FUNCTION_BLOCK FB_Gr00Utility
(*

The function block used to control general utility of the machine.

Constructor: 		Patryk Panylo
Company:		E. Riexinger GmbH
Date:			28.04.2015
Version:			1.00

Date:			Revision:		Who:				Comment
dd.mm.yyyy		x.xx			Initials			comment

*)
VAR_INPUT
	(* Input variables / Eingang Variablen *)
	bSignalStart					:BOOL;						(* Signal "Start" / Signal "Start" *)
	bSignalStop					:BOOL;						(* Signal "Stop" / Signal "Stop" *)
	bSignalAbort					:BOOL;						(* Signal "Abort" / Signal "Abort" *)
	bSignalHome					:BOOL;						(* Signal "Home" / Signal "Grundstellung" *)
	bSignalReference				:BOOL;						(* Signal "Reference" / Signal "Referenz" *)
	bSignalReset					:BOOL;						(* Signal "Reset" / Signal "Reset *)
	bSignalMachinePurge			:BOOL;						(* Machine purge *)
	bAutoStartRelease			:BOOL;						(* Auto start release *)
	bHomeStartRelease			:BOOL;						(* Home start release *)
	bAutoToHome				:BOOL;						(* If auto completed go to home *)
	bHomeCompleted				:BOOL;						(* Home completed signal *)
	bAutoCompleted				:BOOL;						(* Auto completed signal *)
	bAllDoorsClosed 				:BOOL;						(* All doors closed *)
	bAllDoorsLocked 				:BOOL;						(* All doors locked *)
	bLightCurtainOk				:BOOL;						(* Light curtain ok *)
	bExeCounter					:BOOL;						(* Execute counter *)
	bResetCounterUser			:BOOL;						(* Reset counter user *)
	bStartTime					:BOOL;						(* Start measurement of cylce time *)
	bStopTime					:BOOL;						(* Stop measurement of cylce time *)
	bLifetimeOn					:BOOL;						(* Lifetime on *)
	bResetLifetimeAll				:BOOL; 						(* Reset all counters *)
	sLifetimeFilePath				:STRING;					(* File path for life time *)
	sLifetimeFileName			:STRING;					(* File name for life time *)
	bWritePersistent				:BOOL;						(* Write persistent data *)
	bDownTraceDataExe 			:BOOL;						(* Download traceability data *)
	stTraceability					:ST_Traceability;				(* Traceability data *)
	tAdsTimeOut 					:TIME := t#2s;					(* Timout for ads commands *)
END_VAR
VAR_OUTPUT
	(* Output variables / Ausgang Variablen *)
	etMachineMode				:ET_MachineMode;			(* Machine mode *)
	etMachineState				:ET_MachineState;			(* Machine state *)
	bModeAutomatic				:BOOL;						(* Machine mode automatic *)
	bModeHome					:BOOL;						(* Machine mode home *)
	bModeManual				:BOOL;						(* Machine mode manual *)
	bMachineRunning				:BOOL;						(* Machine running *)
	bMachineStandstill			:BOOL;						(* Machine standstill *)
	bMachinePurge				:BOOL;						(* Machine purge *)
	bConfirmAlarm				:BOOL;						(* Alarm confirm *)
	rActOverride					:REAL;						(* Actual override *)
	lrLifetimeAll					:LREAL;						(* Lifetime *)
	lrLifetimeAfterTrunOn			:LREAL;						(* Time after turn on *)
	lrActCycleTime				:LREAL;						(* Actual cycle time *)
	dwCycleTime					:DWORD;					(* Cycletime in 0.01sec / Zykluszeit in 0.01Sekunden *)
END_VAR
VAR_IN_OUT
	(* Input Output variables / Ausgang Variablen *)
	etMachineModeReq			:ET_MachineMode;			(* Machine mode request *)
	rGlobalOverride				:REAL;						(* Global override *)
	udnCounterTotal				:UDINT;						(* Total counter *)
	udnCounterUser				:UDINT;						(* Total counter *)
END_VAR
VAR
	(* Enummerations *)

	(* Variables *)
	nIRHSCtrlCnt					:INT;
	nIRHSZoneCnt				:INT;
	lrIRHSSetpointLeftSide			:LREAL;
	lrIRHSSetpointRightSide		:LREAL;

	bTraceExe					:BOOL;
	ftTraceExe					:F_TRIG;
	rtDownTraceDataExe			:R_TRIG;
	rtDownTraceDataReset		:R_TRIG;
	udnTraceSampleCnt			:UDINT;
	udnTraceDataCnt				:UDINT;

	(* References *)

	(* Interfaces *)

	(* Instances *)
	fbModeSelector				:FB_ModeSelector;			(* Mode selector *)
	fbOverride					:FB_Override;					(* Override *)
	fbLifetime					:FB_TimeHoursCounter;		(* Machine lifetime *)
	fbCounterTotal				:FB_Counter;					(* Counter total *)
	fbCounterUser				:FB_Counter;					(* Counter user *)
	rtResetCounterUser			:R_TRIG;						(* Reset counter user *)
	fbCylceTime					:FB_Timer;					(* Machine cycle time *)
	fbSUPS						:FB_S_UPS_CX51x0;			(*  The function block FB_S_UPS_CX51x0 can be used on CX devices with one-second UPS to control the one-second UPS from the PLC *)
	fbWritePersistentData			:WritePersistentData;			(*  Write Persistent *)
	fbGetCurTaskIdx				:GETCURTASKINDEX;			(* This function block finds the task index of the task from which it is called *)
	fbRTC						:FB_RTC;					(* Get current time *)
	fbTraceability					:FB_Traceability;				(* Traceability *)
	rtMachinePurge				:R_TRIG;
	SystemTaskInfoArr: INT;
END_VAR


A_OperationMode();
A_Override();
A_Counter();
A_CycleTime();
A_MachinePurge();
A_Persistent();
A_PlcTaskSystemInfo();
A_RTC();
A_Traceability();

ACTION A_Counter:

(* Hours counter *)
fbLifetime(
	bEnable := TRUE,
	bDeleteAll := bResetLifetimeAll,
	sAmsNetId := sgAmsNetId,
	bCount := bLifetimeOn,
	bSave := FALSE,
	sFilePath := sLifetimeFilePath,
	sFileName := sLifetimeFileName,
	tSaveIntervall := t#5m,
	tTimeout := tAdsTimeOut,
	lrAllOverHours => lrLifetimeAll,
	lrNoRetainHours => lrLifetimeAfterTrunOn,
 );

(* General counter *)
fbCounterTotal(
	bEnable := TRUE,
	bExecute := bExeCounter,
	bReset := fbCounterTotal.bOverflow,
	udnCounter := udnCounterTotal
);

rtResetCounterUser(CLK:= bResetCounterUser);

fbCounterUser(
	bEnable := TRUE,
	bExecute := bExeCounter,
	bReset := rtResetCounterUser.Q
			 OR fbCounterUser.bOverflow,
	udnCounter := udnCounterUser
);
END_ACTION

ACTION A_CycleTime:

(* Cylce time *)
fbCylceTime(
	bEnable := TRUE,
	bReset := FALSE,
	bStartStop := bStartTime
			        AND bModeAutomatic,
	bStop := bStopTime
		        OR bMachineStandstill,
	tMaxTime := ,
	stRefTime => ,
	stActTime => ,
	stRestTime =>
);

dwCycleTime := fbCylceTime.stActTime.dwDeciSec;
END_ACTION

ACTION A_MachinePurge:

rtMachinePurge(CLK := 	bSignalMachinePurge);

IF NOT bModeAutomatic
     OR bAutoCompleted
THEN
	bMachinePurge := FALSE;

ELSIF rtMachinePurge.Q
THEN
	bMachinePurge := TRUE;
END_IF
END_ACTION

ACTION A_OperationMode:

(* Operation mode control *)
fbModeSelector(
	bStart := bSignalStart,
	bStop := bSignalStop,
	bAbort := bSignalAbort,
	bHome := bSignalHome,
	bReset := bSignalReset,
	bReference := bSignalReference,
	bAutoStartRelease := bAutoStartRelease,
	bHomeStartRelease := bHomeStartRelease,
	bAutoToHome := bAutoToHome,
	bHomeCompleted := bHomeCompleted,
	bAutoCompleted := bAutoCompleted,
	bAllDoorsClosed  := bAllDoorsClosed,
	bAllDoorsLocked := bAllDoorsLocked,
	bLightCurtainOk := bLightCurtainOk,
	etMachineMode => etMachineMode,
	etMachineState => etMachineState,
	bModeAutomatic => bModeAutomatic,
	bModeHome => bModeHome,
	bModeManual => bModeManual,
	bMachineRunning => bMachineRunning,
	bMachineStandstill => bMachineStandstill,
	bConfirmAlarm => bConfirmAlarm,
	etMachineModeReq := etMachineModeReq
);
END_ACTION

ACTION A_Override:

(* Override control *)
fbOverride(
	bEnable := TRUE,
	bBypassAccDec := bModeManual,
	bSetOverideMax := bModeAutomatic,
	rAcc := rgGr00AdsOverrideAcc,
	rDec := rgGr01AdsOverrideDec,
	rSetOverride := rGlobalOverride,
	rActOverride => rActOverride
);
END_ACTION

ACTION A_Persistent:

(*  The function block FB_S_UPS_CX51x0 can be used on CX devices with one-second UPS to control the one-second UPS from the PLC *)
fbSUPS(
	sNetID := sgAmsNetId,													(* AmsNetID of the controller. *)
	iPLCPort := AMSPORT_R0_PLC_RTS1,									(* Port number of the PLC runtime system (AMSPORT_R0_PLC_RTS1 = 801, AMSPORT_R0_PLC_RTS2 = 811, AMSPORT_R0_PLC_RTS3 = 821, AMSPORT_R0_PLC_RTS4 = 831). *)
	iUPSPort := 16#588,													(* Port number via which the UPS status is read (standard value is 16#588) *)
	tTimeout := DEFAULT_ADS_TIMEOUT,									(* ADS Timeout *)
	eUpsMode := eSUPS_WrPersistData_Shutdown,							(* The eUpsMode defines whether persistent data are to be written and whether a QuickShutdown is to be performed.
																		Standard value is eSUPS_WrPersistData_Shutdown, i.e. with writing of the persistent data and then QuickShutdown. See E_S_UPS_Mode. *)
	ePersistentMode := SPDM_2PASS,										(* Mode for the writing of the persistent data. Standard value is SPDM_2PASS *)
	tRecoverTime := t#10s													(* Time after which the UPS reverts to the PowerOK status in the case of UPS modes without shutdown.
																	   	    The tRecoverTime must be somewhat longer than the maximum holding time of the UPS, since the UPS switches off even when the voltage returns. *)
);


(* If persistent variables are defined in one of the PLC's runtime systems, then their current values are stored in a file in the TwinCAT\Boot directory when the TwinCAT system stops (after the last PLC cycle). *)
fbWritePersistentData(
	NETID := sgAmsNetId,
	PORT := AMSPORT_R0_PLC_RTS1,
	START := bWritePersistent
			   AND NOT fbWritePersistentData.BUSY,
	TMOUT := DEFAULT_ADS_TIMEOUT
);
END_ACTION

ACTION A_PlcTaskSystemInfo:

fbGetCurTaskIdx();

// lrActCycleTime := UDINT_TO_LREAL(SystemTaskInfoArr[fbGetCurTaskIdx.index].cycleTime) / 10000000;




fbGetCurTaskIdx();

GVL._PlcTaskSystemInfo := _TaskInfo[fbGetCurTaskIdx.index];

lrActCycleTime := UDINT_TO_LREAL(_TaskInfo[fbGetCurTaskIdx.index].CycleTime) / 10000000;
END_ACTION

ACTION A_RTC:

fbRTC(
	stDateTime => stgGr00DateTime
);
END_ACTION

ACTION A_Traceability:

stTraceability.sDateTime := stgGr00DateTime.sDateTime;

stTraceability.stSettings.sPath := sTracePath(*CONCAT(CONCAT(sTracePath,fbRTC.sDate),'\')*);
stTraceability.stSettings.sFileName := stgGr00DateTime.sDateTime;
stTraceability.stSettings.sFileExtension := sTraceFileExtension;

rtDownTraceDataReset(
	CLK := bModeAutomatic
);

IF rtDownTraceDataReset.Q
THEN
	udnTraceSampleCnt := 0;
	MEMSET(ADR(stTraceability.arstData), 0, SIZEOF(stTraceability.arstData));
END_IF

rtDownTraceDataExe(
	CLK := bTraceEnable
		    AND bDownTraceDataExe
);

IF rtDownTraceDataExe.Q
     AND udnTraceSampleCnt < udnTraceSampleMax
THEN
	udnTraceDataCnt := 0;
	udnTraceSampleCnt := udnTraceSampleCnt +1;
	(*1*)
	udnTraceDataCnt := udnTraceDataCnt + 1;
	stTraceability.arstData[udnTraceSampleCnt,udnTraceDataCnt].sName := 'Time';
	stTraceability.arstData[udnTraceSampleCnt,udnTraceDataCnt].sValue := stgGr00DateTime.sDateTime;
	stTraceability.arstData[udnTraceSampleCnt,udnTraceDataCnt].sUnit := '';

	(*2*)
	udnTraceDataCnt := udnTraceDataCnt + 1;
	stTraceability.arstData[udnTraceSampleCnt,udnTraceDataCnt].sName := 'Cntr';
	stTraceability.arstData[udnTraceSampleCnt,udnTraceDataCnt].sValue := UDINT_TO_STRING(stgGr00HMI.stPLCTOHMI.udnCounterTotal);
	stTraceability.arstData[udnTraceSampleCnt,udnTraceDataCnt].sUnit := '';

END_IF

(*ftTraceExe(CLK := bgGr00ModeAutomatic);*)
fbTraceability(
	bEnable := bTraceEnable,
	bExecute := bAutoCompleted
			     (*OR
			     (NOT bAutoCompleted
			      AND (bSignalStop OR bSignalAbort)
			      AND ftTraceExe.Q)*)
			     OR bTraceExe,
	stTraceability := stTraceability
);
END_ACTION

END_FUNCTION_BLOCK

(* stored: Version 1.1.0.1, ProductVersion 3.1.4024.15
   POU FB_Gr00Utility: Id {2dde8993-b0f9-4f82-b192-aa7b8cf4d050}, SpecialFunc None
   Action A_Counter: Id {a76de720-a836-4d60-a585-108dc094c4d1}
   Action A_CycleTime: Id {be029e3a-8ddb-4b33-be5e-5d356f1a1ee0}
   Action A_MachinePurge: Id {0ab65900-954c-49a1-971b-74fc5e33a980}
   Action A_OperationMode: Id {42a518b3-dd1b-4820-a289-1209514f9c62}
   Action A_Override: Id {78915dc2-c243-4cf7-ba34-72ce962f01f1}
   Action A_Persistent: Id {fa4aa848-7ac9-4ab5-b018-4f0e657e5d2b}
   Action A_PlcTaskSystemInfo: Id {3de26191-b8ed-43bc-8322-92490ef8f70b}
   Action A_RTC: Id {6cec8227-c097-4090-bb19-8d819d2ab91a}
   Action A_Traceability: Id {877129ff-9ebe-428b-a868-1b958abf19ee} *)
